(* IEC 61131-3 sources: kkh_knowHow_dgtt/tools/fmse/plc_lib, 31 files *)

(* ---- TYPES.st ---- *)
(*==================================================================================================================
  TYPES  -  enumerations and global constants of the FMSE device FB library
  ----------------------------------------------------------------------------------------------------------------
  Library   : FMSE device FB library (item 10A)              Version : 1.0.0 (2026-11-15)
  Rule      : tools/fmse/examples/item10a_examples.json  _rules.common, decisions D1 - D4
  Purpose   : one place for the state numbers (PackML item 5, device FBs), alarm classes and the time base.
              Load this file FIRST. Enumerations are used qualified (E_DriveState.FAULT); in CODESYS add
              the pragma attribute 'qualified_only', in TIA Portal use INT constants with the same values.
  Timing    : GC_CYCLE_MS = time base of the call counters of every FB. 100 = test bench (one call per
              100 ms tick). In the 10 ms main task set 10 - every time in ms stays the same.
  NOTICE    : ALL VALUES ARE EXAMPLES. Real PLC code is written, reviewed, tested and signed off by qualified
              people. Safety functions only in the F-program.
==================================================================================================================*)
TYPE
  E_AlarmClass : (NONE := 0, A := 1, B := 2, C := 3) INT;          (* decision D3 *)
  E_Reaction : (NONE := 0, ABORT := 1, HOLD := 2, WARNING := 3) INT;
  E_AlarmEvent : (NONE := 0, RAISE := 1, CLEAR := 2) INT;
  E_PackMLState : (UNDEFINED := 0, CLEARING := 1, STOPPED := 2, STARTING := 3, IDLE := 4, SUSPENDED := 5,
                   EXECUTE := 6, STOPPING := 7, ABORTING := 8, ABORTED := 9, HOLDING := 10, HELD := 11,
                   UNHOLDING := 12, SUSPENDING := 13, UNSUSPENDING := 14, RESETTING := 15, COMPLETING := 16,
                   COMPLETE := 17) INT;                             (* item 5, PackML / ISA-TR88 *)
  E_PackMLCmd : (NONE := 0, RESET := 1, START := 2, STOP := 3, HOLD := 4, UNHOLD := 5, SUSPEND := 6,
                 UNSUSPEND := 7, ABORT := 8, CLEAR := 9) INT;
  E_Mode : (UNDEFINED := 0, PRODUCTION := 1, MAINTENANCE := 2, MANUAL := 3) INT;
  E_DriveState : (NOT_READY := 0, READY := 1, RUNNING := 2, FAULT := 9) INT;
  E_MotorState : (STOPPED := 0, STARTING := 1, RUNNING := 2, STOPPING := 3, FAULT := 9) INT;
  E_HsStep : (IDLE := 0, REQUEST := 10, BUSY := 20, DONE := 30) INT;
  E_Quality : (GOOD := 0, UNCERTAIN := 1, BAD := 2) INT;             (* NAMUR NE 43 *)
  E_AiStatus : (OK := 0, FAULT_LOW := 1, UNDER_RANGE := 2, OVER_RANGE := 3, FAULT_HIGH := 4) INT;
END_TYPE

VAR_GLOBAL CONSTANT
  GC_CYCLE_MS : DINT := 100;                  (* time base of the call counters [ms] *)
  GC_N_MAX : DINT := 1000000;                 (* counters stop here (no overflow, 27 h at 100 ms) *)
  GC_BLINK_HALF_MS : DINT := 500;             (* half period of the 1 Hz blink [ms] *)
  GC_LIB_VERSION : WORD := 16#0100;           (* library version 1.0.0 *)
END_VAR

(* ---- F_CmdAllowed.st ---- *)
(*==================================================================================================================
  F_CmdAllowed  -  PackML command allowed in this state and mode? (item 5 tables)
  ----------------------------------------------------------------------------------------------------------------
  Library   : FMSE device FB library (item 10A)              Version : 1.0.0 (2026-11-15)
  Rule      : tools/fmse/examples/item10a_examples.json  _rules.FB_CmdIf
  Purpose   : TRUE when the command is in the mode table (1 Production: all 9, 2 Maintenance: without
              Suspend/Unsuspend, 3 Manual: Reset, Start, Stop, Abort, Clear) AND it is a transition of the
              state model: EDGES with the command label, Stop from every state except Stopped / Stopping /
              Aborting / Aborted / Clearing, Abort from every state except Aborting / Aborted.
  Interface :
    dir  name                type          default   meaning
    IN   iCmd                INT           -         command 1 Reset .. 9 Clear
    IN   iState              INT           -         PackML state 1 .. 17
    IN   iMode               INT           -         1 Production, 2 Maintenance, 3 Manual
  Alarms    : iAlarm = local code a ; Admin.AlarmNo = M*1000 + 10*i + a (decision D2), class per module (D3)
    none
  Timing    : Times are counted in calls: n * GC_CYCLE_MS >= t_ms (GC_CYCLE_MS = 100 ms = test bench, TYPES.st).
              In the 10 ms main task set GC_CYCLE_MS := 10 (same behaviour, 10 ms resolution) or replace a counter
              by a TON: ton(IN := <condition>, PT := T#2s); IF ton.Q THEN ... (one call later than the counter).
  Siemens   : SCL (TIA Portal): the same statements; local names are written with '#' (#xRst), the VAR section is
              VAR (STAT) of an FB with an instance DB, R_TRIG / TON are multi-instances, enumerations become INT
              constants (E_DriveState.FAULT -> 9), MIN / LIMIT exist, '16#0080' is written W#16#80 for a WORD.
  NOTICE    : ALL VALUES ARE EXAMPLES. Real PLC code is written, reviewed, tested and signed off by qualified
              people. Safety functions only in the F-program; this FB only reads F-copies and writes no F-signal.
==================================================================================================================*)
FUNCTION F_CmdAllowed : BOOL
VAR_INPUT  (* signals *)
  iCmd : INT;                               (* command 1 Reset .. 9 Clear *)
  iState : INT;                             (* PackML state 1 .. 17 *)
  iMode : INT;                              (* 1 Production, 2 Maintenance, 3 Manual *)
END_VAR
VAR  (* internal *)
  xInMode : BOOL;                           (* command allowed in the mode *)
END_VAR
F_CmdAllowed := FALSE;
CASE iMode OF
  E_Mode.PRODUCTION:
    xInMode := iCmd >= E_PackMLCmd.RESET AND iCmd <= E_PackMLCmd.CLEAR;
  E_Mode.MAINTENANCE:
    xInMode := (iCmd >= E_PackMLCmd.RESET AND iCmd <= E_PackMLCmd.UNHOLD) OR iCmd = E_PackMLCmd.ABORT
               OR iCmd = E_PackMLCmd.CLEAR;
  E_Mode.MANUAL:
    xInMode := (iCmd >= E_PackMLCmd.RESET AND iCmd <= E_PackMLCmd.STOP) OR iCmd = E_PackMLCmd.ABORT
               OR iCmd = E_PackMLCmd.CLEAR;
ELSE
  xInMode := FALSE;
END_CASE
IF NOT xInMode OR iState < E_PackMLState.CLEARING OR iState > E_PackMLState.COMPLETE THEN
  RETURN;
END_IF
CASE iCmd OF
  E_PackMLCmd.RESET:
    F_CmdAllowed := iState = E_PackMLState.STOPPED OR iState = E_PackMLState.COMPLETE;
  E_PackMLCmd.START:
    F_CmdAllowed := iState = E_PackMLState.IDLE;
  E_PackMLCmd.STOP:
    CASE iState OF
      E_PackMLState.CLEARING, E_PackMLState.STOPPED, E_PackMLState.STOPPING..E_PackMLState.ABORTED:
        F_CmdAllowed := FALSE;
    ELSE
      F_CmdAllowed := TRUE;
    END_CASE
  E_PackMLCmd.HOLD, E_PackMLCmd.SUSPEND:
    F_CmdAllowed := iState = E_PackMLState.EXECUTE;
  E_PackMLCmd.UNHOLD:
    F_CmdAllowed := iState = E_PackMLState.HELD;
  E_PackMLCmd.UNSUSPEND:
    F_CmdAllowed := iState = E_PackMLState.SUSPENDED;
  E_PackMLCmd.ABORT:
    F_CmdAllowed := iState <> E_PackMLState.ABORTING AND iState <> E_PackMLState.ABORTED;
  E_PackMLCmd.CLEAR:
    F_CmdAllowed := iState = E_PackMLState.ABORTED;
END_CASE
END_FUNCTION

(* ---- FB_AlarmMgr.st ---- *)
(*==================================================================================================================
  FB_AlarmMgr  -  module alarm manager: AlarmNo, WarningNo, class, reaction (D2 + D3)
  ----------------------------------------------------------------------------------------------------------------
  Library   : FMSE device FB library (item 10A)              Version : 1.0.0 (2026-11-15)
  Rule      : tools/fmse/examples/item10a_examples.json  _rules.alarm_manager
  Purpose   : Called once per alarm change (iEvent 1 = on, 2 = off; 0 = only evaluate) with the instance i, the
              local code a and the class of that alarm (class table generated from the library, item 10B).
              Admin.AlarmNo = best active class A/B alarm (A before B, earlier before later), Admin.WarningNo =
              earliest active class C, iAlarmClass for FB_SignalTower, iReaction for the PackML core.
  Interface :
    dir  name                type          default   meaning
    IN   iEvent              INT           -         0 none, 1 alarm on, 2 alarm off
    IN   iInst               INT           -         instance number i (0 = module level)
    IN   iCode               INT           -         local alarm code a (1 .. 9)
    IN   iClass              INT           -         class 1 A, 2 B, 3 C
    CFG  iModule             INT           2         module number M (M02 -> 2)
    OUT  iAlarmNo            INT           -         Admin.AlarmNo = M*1000 + 10*i + a
    OUT  iWarningNo          INT           -         Admin.WarningNo
    OUT  iAlarmClass         INT           -         0 none, 1 A, 2 B, 3 C
    OUT  iReaction           INT           -         0 none, 1 Abort, 2 Hold if Execute, 3 warning
    OUT  iActive             INT           -         number of active alarms
    OUT  xOverflow           BOOL          -         active list full
  Alarms    : iAlarm = local code a ; Admin.AlarmNo = M*1000 + 10*i + a (decision D2), class per module (D3)
    none
  Timing    : Times are counted in calls: n * GC_CYCLE_MS >= t_ms (GC_CYCLE_MS = 100 ms = test bench, TYPES.st).
              In the 10 ms main task set GC_CYCLE_MS := 10 (same behaviour, 10 ms resolution) or replace a counter
              by a TON: ton(IN := <condition>, PT := T#2s); IF ton.Q THEN ... (one call later than the counter).
  Siemens   : SCL (TIA Portal): the same statements; local names are written with '#' (#xRst), the VAR section is
              VAR (STAT) of an FB with an instance DB, R_TRIG / TON are multi-instances, enumerations become INT
              constants (E_DriveState.FAULT -> 9), MIN / LIMIT exist, '16#0080' is written W#16#80 for a WORD.
  NOTICE    : ALL VALUES ARE EXAMPLES. Real PLC code is written, reviewed, tested and signed off by qualified
              people. Safety functions only in the F-program; this FB only reads F-copies and writes no F-signal.
==================================================================================================================*)
FUNCTION_BLOCK FB_AlarmMgr
VAR_INPUT  (* signals *)
  iEvent : INT;                             (* 0 none, 1 alarm on, 2 alarm off *)
  iInst : INT;                              (* instance number i (0 = module level) *)
  iCode : INT;                              (* local alarm code a (1 .. 9) *)
  iClass : INT;                             (* class 1 A, 2 B, 3 C *)
END_VAR
VAR_INPUT  (* configuration (set once, defaults = example values) *)
  iModule : INT := 2;                       (* module number M (M02 -> 2) *)
END_VAR
VAR_OUTPUT  (* outputs *)
  iAlarmNo : INT;                           (* Admin.AlarmNo = M*1000 + 10*i + a *)
  iWarningNo : INT;                         (* Admin.WarningNo *)
  iAlarmClass : INT;                        (* 0 none, 1 A, 2 B, 3 C *)
  iReaction : INT;                          (* 0 none, 1 Abort, 2 Hold if Execute, 3 warning *)
  iActive : INT;                            (* number of active alarms *)
  xOverflow : BOOL;                         (* active list full *)
END_VAR
VAR CONSTANT  (* constants *)
  MAX_ACT : INT := 32;                      (* size of the active list *)
END_VAR
VAR  (* internal *)
  aiNo : ARRAY[1..MAX_ACT] OF INT;          (* active alarm numbers (0 = free) *)
  aiCls : ARRAY[1..MAX_ACT] OF INT;         (* class of each active alarm *)
  adiOrd : ARRAY[1..MAX_ACT] OF DINT;       (* activation order *)
  diOrder : DINT;                           (* activation counter *)
  iNo : INT;                                (* number of this event *)
  k : INT;                                  (* loop index *)
  iFound : INT;                             (* slot of iNo (0 = not active) *)
  iFree : INT;                              (* first free slot *)
  iBest : INT;                              (* slot of the best A/B alarm *)
  iBestW : INT;                             (* slot of the earliest warning *)
END_VAR
IF iEvent <> E_AlarmEvent.NONE THEN
  iNo := iModule * 1000 + 10 * iInst + iCode;
  iFound := 0;
  iFree := 0;
  FOR k := 1 TO MAX_ACT DO
    IF aiNo[k] = iNo AND iFound = 0 THEN
      iFound := k;
    END_IF
    IF aiNo[k] = 0 AND iFree = 0 THEN
      iFree := k;
    END_IF
  END_FOR
  IF iEvent = E_AlarmEvent.RAISE AND iFound = 0 THEN
    IF iFree > 0 THEN
      diOrder := diOrder + 1;
      aiNo[iFree] := iNo;
      aiCls[iFree] := iClass;
      adiOrd[iFree] := diOrder;
    ELSE
      xOverflow := TRUE;
    END_IF
  ELSIF iEvent = E_AlarmEvent.CLEAR AND iFound > 0 THEN
    aiNo[iFound] := 0;
    aiCls[iFound] := 0;
    adiOrd[iFound] := 0;
  END_IF
END_IF
(* evaluate: best class A/B alarm by (class, activation order), earliest class C warning *)
iBest := 0;
iBestW := 0;
iActive := 0;
FOR k := 1 TO MAX_ACT DO
  IF aiNo[k] <> 0 THEN
    iActive := iActive + 1;
    IF aiCls[k] = E_AlarmClass.A OR aiCls[k] = E_AlarmClass.B THEN
      IF iBest = 0 THEN
        iBest := k;
      ELSIF aiCls[k] < aiCls[iBest] OR (aiCls[k] = aiCls[iBest] AND adiOrd[k] < adiOrd[iBest]) THEN
        iBest := k;
      END_IF
    ELSIF aiCls[k] = E_AlarmClass.C THEN
      IF iBestW = 0 THEN
        iBestW := k;
      ELSIF adiOrd[k] < adiOrd[iBestW] THEN
        iBestW := k;
      END_IF
    END_IF
  END_IF
END_FOR
IF iBest > 0 THEN
  iAlarmNo := aiNo[iBest];
  iAlarmClass := aiCls[iBest];
ELSE
  iAlarmNo := 0;
  IF iBestW > 0 THEN
    iAlarmClass := E_AlarmClass.C;
  ELSE
    iAlarmClass := E_AlarmClass.NONE;
  END_IF
END_IF
IF iBestW > 0 THEN
  iWarningNo := aiNo[iBestW];
ELSE
  iWarningNo := 0;
END_IF
CASE iAlarmClass OF
  E_AlarmClass.A: iReaction := E_Reaction.ABORT;
  E_AlarmClass.B: iReaction := E_Reaction.HOLD;
  E_AlarmClass.C: iReaction := E_Reaction.WARNING;
ELSE
  iReaction := E_Reaction.NONE;
END_CASE
END_FUNCTION_BLOCK

(* ---- FB_AnalogIn.st ---- *)
(*==================================================================================================================
  FB_AnalogIn  -  4-20 mA analog input: scaling, NAMUR NE 43 quality, substitute value (item 9)
  ----------------------------------------------------------------------------------------------------------------
  Library   : FMSE device FB library (item 10A)              Version : 1.0.0 (2026-11-15)
  Rule      : tools/fmse/examples/item10a_examples.json  item9_examples.json _rules.analog
  Codegen   : item 8 pattern ANALOG_P, ANALOG_T -> st_codegen.py calls this FB (x<Signal> / q<Signal>)
  Purpose   : raw 0..27648 = 4..20 mA (Siemens-style card scaling - check yours). NE 43: <= 3.6 mA BAD (wire
              break), < 3.8 UNCERTAIN, <= 20.5 GOOD, < 21.0 UNCERTAIN, else BAD. rValue = clamped value for
              GOOD / UNCERTAIN, substitute rLo for BAD (the module must not use a BAD value).
  Interface :
    dir  name                type          default   meaning
    IN   iValue              INT           -         raw value of the card (AI)
    CFG  rLo                 REAL          0.0       value at 4 mA
    CFG  rHi                 REAL          10.0      value at 20 mA
    OUT  rMa                 REAL          -         current [mA]
    OUT  rValueLin           REAL          -         linear value (not clamped)
    OUT  rValue              REAL          -         value to use (clamped / substitute)
    OUT  iQuality            INT           -         0 GOOD, 1 UNCERTAIN, 2 BAD
    OUT  iStatus             INT           -         0 ok, 1 fault low, 2 under, 3 over, 4 fault high
    OUT  xGood               BOOL          -         quality GOOD
    OUT  iAlarm              INT           -         local alarm code (0 = none)
  Alarms    : iAlarm = local code a ; Admin.AlarmNo = M*1000 + 10*i + a (decision D2), class per module (D3)
    3  signal quality bad/uncertain (NAMUR NE 43)
  Timing    : Times are counted in calls: n * GC_CYCLE_MS >= t_ms (GC_CYCLE_MS = 100 ms = test bench, TYPES.st).
              In the 10 ms main task set GC_CYCLE_MS := 10 (same behaviour, 10 ms resolution) or replace a counter
              by a TON: ton(IN := <condition>, PT := T#2s); IF ton.Q THEN ... (one call later than the counter).
  Siemens   : SCL (TIA Portal): the same statements; local names are written with '#' (#xRst), the VAR section is
              VAR (STAT) of an FB with an instance DB, R_TRIG / TON are multi-instances, enumerations become INT
              constants (E_DriveState.FAULT -> 9), MIN / LIMIT exist, '16#0080' is written W#16#80 for a WORD.
  NOTICE    : ALL VALUES ARE EXAMPLES. Real PLC code is written, reviewed, tested and signed off by qualified
              people. Safety functions only in the F-program; this FB only reads F-copies and writes no F-signal.
==================================================================================================================*)
FUNCTION_BLOCK FB_AnalogIn
VAR_INPUT  (* signals *)
  iValue : INT;                             (* raw value of the card (AI) *)
END_VAR
VAR_INPUT  (* configuration (set once, defaults = example values) *)
  rLo : REAL := 0.0;                        (* value at 4 mA *)
  rHi : REAL := 10.0;                       (* value at 20 mA *)
END_VAR
VAR_OUTPUT  (* outputs *)
  rMa : REAL;                               (* current [mA] *)
  rValueLin : REAL;                         (* linear value (not clamped) *)
  rValue : REAL;                            (* value to use (clamped / substitute) *)
  iQuality : INT;                           (* 0 GOOD, 1 UNCERTAIN, 2 BAD *)
  iStatus : INT;                            (* 0 ok, 1 fault low, 2 under, 3 over, 4 fault high *)
  xGood : BOOL;                             (* quality GOOD *)
  iAlarm : INT;                             (* local alarm code (0 = none) *)
END_VAR
rMa := 4.0 + 16.0 * INT_TO_REAL(iValue) / 27648.0;
IF rMa <= 3.6 THEN
  iQuality := E_Quality.BAD;
  iStatus := E_AiStatus.FAULT_LOW;            (* wire break *)
ELSIF rMa < 3.8 THEN
  iQuality := E_Quality.UNCERTAIN;
  iStatus := E_AiStatus.UNDER_RANGE;
ELSIF rMa <= 20.5 THEN
  iQuality := E_Quality.GOOD;
  iStatus := E_AiStatus.OK;
ELSIF rMa < 21.0 THEN
  iQuality := E_Quality.UNCERTAIN;
  iStatus := E_AiStatus.OVER_RANGE;
ELSE
  iQuality := E_Quality.BAD;
  iStatus := E_AiStatus.FAULT_HIGH;
END_IF
rValueLin := rLo + (rHi - rLo) * (rMa - 4.0) / 16.0;
IF iQuality = E_Quality.BAD THEN
  rValue := rLo;                              (* substitute value *)
ELSE
  rValue := LIMIT(rLo, rValueLin, rHi);
END_IF
xGood := iQuality = E_Quality.GOOD;
IF xGood THEN
  iAlarm := 0;
ELSE
  iAlarm := 3;                                (* signal quality bad / uncertain *)
END_IF
END_FUNCTION_BLOCK

(* ---- FB_CmdIf.st ---- *)
(*==================================================================================================================
  FB_CmdIf  -  command interface of the module data block (4-phase echo, decision D1)
  ----------------------------------------------------------------------------------------------------------------
  Library   : FMSE device FB library (item 10A)              Version : 1.0.0 (2026-11-15)
  Rule      : tools/fmse/examples/item10a_examples.json  _rules.FB_CmdIf
  Purpose   : The cell controller writes CntrlCmd + sets CmdChangeRequest in ONE FC16 write. On the rising edge
              the module evaluates the command (F_CmdAllowed) -> CmdAck (Status.Bits bit8, iCmdExec one call
              for the PackML core) or CmdRej (bit9; the module sets Admin.WarningNo = M*1000 + 900 + command).
              The CC clears the request, then the module clears the echo. One writer per word, no command twice.
  Interface :
    dir  name                type          default   meaning
    IN   iCntrlCmd           INT           -         data block word CntrlCmd (written by the CC)
    IN   xCmdChangeRequest   BOOL          -         word 3 bit0 (written by the CC)
    IN   iState              INT           2         PackML state of the module
    IN   iMode               INT           1         mode of the module
    OUT  xCmdAck             BOOL          -         echo: accepted (Status.Bits bit8)
    OUT  xCmdRej             BOOL          -         echo: rejected (Status.Bits bit9)
    OUT  iCmdExec            INT           -         command to execute, one call (0 = none)
    OUT  iLastCmd            INT           -         last evaluated command
    OUT  iRejectCount        INT           -         rejected commands
  Alarms    : iAlarm = local code a ; Admin.AlarmNo = M*1000 + 10*i + a (decision D2), class per module (D3)
    none
  Timing    : Times are counted in calls: n * GC_CYCLE_MS >= t_ms (GC_CYCLE_MS = 100 ms = test bench, TYPES.st).
              In the 10 ms main task set GC_CYCLE_MS := 10 (same behaviour, 10 ms resolution) or replace a counter
              by a TON: ton(IN := <condition>, PT := T#2s); IF ton.Q THEN ... (one call later than the counter).
  Siemens   : SCL (TIA Portal): the same statements; local names are written with '#' (#xRst), the VAR section is
              VAR (STAT) of an FB with an instance DB, R_TRIG / TON are multi-instances, enumerations become INT
              constants (E_DriveState.FAULT -> 9), MIN / LIMIT exist, '16#0080' is written W#16#80 for a WORD.
  NOTICE    : ALL VALUES ARE EXAMPLES. Real PLC code is written, reviewed, tested and signed off by qualified
              people. Safety functions only in the F-program; this FB only reads F-copies and writes no F-signal.
==================================================================================================================*)
FUNCTION_BLOCK FB_CmdIf
VAR_INPUT  (* signals *)
  iCntrlCmd : INT;                          (* data block word CntrlCmd (written by the CC) *)
  xCmdChangeRequest : BOOL;                 (* word 3 bit0 (written by the CC) *)
  iState : INT := 2;                        (* PackML state of the module *)
  iMode : INT := 1;                         (* mode of the module *)
END_VAR
VAR_OUTPUT  (* outputs *)
  xCmdAck : BOOL;                           (* echo: accepted (Status.Bits bit8) *)
  xCmdRej : BOOL;                           (* echo: rejected (Status.Bits bit9) *)
  iCmdExec : INT;                           (* command to execute, one call (0 = none) *)
  iLastCmd : INT;                           (* last evaluated command *)
  iRejectCount : INT;                       (* rejected commands *)
END_VAR
VAR  (* internal *)
  rtReq : R_TRIG;                           (* edge of xCmdChangeRequest *)
END_VAR
rtReq(CLK := xCmdChangeRequest);
iCmdExec := 0;
IF rtReq.Q THEN
  iLastCmd := iCntrlCmd;
  IF F_CmdAllowed(iCmd := iCntrlCmd, iState := iState, iMode := iMode) THEN
    xCmdAck := TRUE;
    iCmdExec := iCntrlCmd;
  ELSE
    xCmdRej := TRUE;
    iRejectCount := iRejectCount + 1;
  END_IF
END_IF
IF NOT xCmdChangeRequest THEN                 (* phase 4: the CC has cleared the request *)
  xCmdAck := FALSE;
  xCmdRej := FALSE;
END_IF
END_FUNCTION_BLOCK

(* ---- FB_ContactorPair.st ---- *)
(*==================================================================================================================
  FB_ContactorPair  -  redundant contactor pair with EDM
  ----------------------------------------------------------------------------------------------------------------
  Library   : FMSE device FB library (item 10A)              Version : 1.0.0 (2026-11-15)
  Rule      : tools/fmse/examples/item10a_examples.json  _rules.fb_library (= FB_Edm, bInverted TRUE)
  Codegen   : item 8 pattern CONT_PAIR_EDM -> st_codegen.py calls this FB (x<Signal> / q<Signal>)
  Purpose   : Wrapper of FB_Edm with bInverted TRUE. The F-output Enable is written only by the F-program;
              xCmd is its read-only F-copy.
  Interface :
    dir  name                type          default   meaning
    IN   xCmd                BOOL          -         F-copy of the F-output Enable
    IN   xEDM                BOOL          TRUE      NC mirror contacts in series (DI), TRUE = open
    IN   xReset              BOOL          -         fault reset, rising edge
    CFG  tEdm_ms             DINT          300       feedback time [ms]
    OUT  xOn                 BOOL          -         output on and feedback ok
    OUT  xError              BOOL          -         error latched (see alarms)
    OUT  iAlarm              INT           -         local alarm code (0 = none)
  Alarms    : iAlarm = local code a ; Admin.AlarmNo = M*1000 + 10*i + a (decision D2), class per module (D3)
    1  feedback does not follow (welded / not switching)
  Timing    : Times are counted in calls: n * GC_CYCLE_MS >= t_ms (GC_CYCLE_MS = 100 ms = test bench, TYPES.st).
              In the 10 ms main task set GC_CYCLE_MS := 10 (same behaviour, 10 ms resolution) or replace a counter
              by a TON: ton(IN := <condition>, PT := T#2s); IF ton.Q THEN ... (one call later than the counter).
  Siemens   : SCL (TIA Portal): the same statements; local names are written with '#' (#xRst), the VAR section is
              VAR (STAT) of an FB with an instance DB, R_TRIG / TON are multi-instances, enumerations become INT
              constants (E_DriveState.FAULT -> 9), MIN / LIMIT exist, '16#0080' is written W#16#80 for a WORD.
  NOTICE    : ALL VALUES ARE EXAMPLES. Real PLC code is written, reviewed, tested and signed off by qualified
              people. Safety functions only in the F-program; this FB only reads F-copies and writes no F-signal.
==================================================================================================================*)
FUNCTION_BLOCK FB_ContactorPair
VAR_INPUT  (* signals *)
  xCmd : BOOL;                              (* F-copy of the F-output Enable *)
  xEDM : BOOL := TRUE;                      (* NC mirror contacts in series (DI), TRUE = open *)
  xReset : BOOL;                            (* fault reset, rising edge *)
END_VAR
VAR_INPUT  (* configuration (set once, defaults = example values) *)
  tEdm_ms : DINT := 300;                    (* feedback time [ms] *)
END_VAR
VAR_OUTPUT  (* outputs *)
  xOn : BOOL;                               (* output on and feedback ok *)
  xError : BOOL;                            (* error latched (see alarms) *)
  iAlarm : INT;                             (* local alarm code (0 = none) *)
END_VAR
VAR  (* internal *)
  fbEdm : FB_Edm;                           (* EDM *)
END_VAR
fbEdm(xCmd := xCmd, xFb := xEDM, xReset := xReset, tEdm_ms := tEdm_ms, bInverted := TRUE);
xOn := fbEdm.xOn;
xError := fbEdm.xError;
iAlarm := fbEdm.iAlarm;
END_FUNCTION_BLOCK

(* ---- FB_Door2Ch.st ---- *)
(*==================================================================================================================
  FB_Door2Ch  -  guard door switch (2 channels, no locking)
  ----------------------------------------------------------------------------------------------------------------
  Library   : FMSE device FB library (item 10A)              Version : 1.0.0 (2026-11-15)
  Rule      : tools/fmse/examples/item10a_examples.json  _rules.fb_library (= FB_Safe2Ch)
  Codegen   : item 8 pattern DOOR_2CH -> st_codegen.py calls this FB (x<Signal> / q<Signal>)
  Purpose   : Wrapper with the item-8 signal names: xClosed / xClosed2 -> FB_Safe2Ch xCh1 / xCh2.
              Diagnosis and HMI only - the safety function is in the F-program.
  Interface :
    dir  name                type          default   meaning
    IN   xClosed             BOOL          -         door closed channel 1 F-copy
    IN   xClosed2            BOOL          -         door closed channel 2 F-copy
    IN   xReset              BOOL          -         fault reset, rising edge
    CFG  tDisc_ms            DINT          500       discrepancy time [ms]
    OUT  xSafe               BOOL          -         closed / free and reset (FB_Safe2Ch.xOk)
    OUT  xResetReq           BOOL          -         waiting for a reset
    OUT  xDiscErr            BOOL          -         discrepancy latched
    OUT  iAlarm              INT           -         local alarm code (0 = none)
  Alarms    : iAlarm = local code a ; Admin.AlarmNo = M*1000 + 10*i + a (decision D2), class per module (D3)
    1  discrepancy
  Timing    : Times are counted in calls: n * GC_CYCLE_MS >= t_ms (GC_CYCLE_MS = 100 ms = test bench, TYPES.st).
              In the 10 ms main task set GC_CYCLE_MS := 10 (same behaviour, 10 ms resolution) or replace a counter
              by a TON: ton(IN := <condition>, PT := T#2s); IF ton.Q THEN ... (one call later than the counter).
  Siemens   : SCL (TIA Portal): the same statements; local names are written with '#' (#xRst), the VAR section is
              VAR (STAT) of an FB with an instance DB, R_TRIG / TON are multi-instances, enumerations become INT
              constants (E_DriveState.FAULT -> 9), MIN / LIMIT exist, '16#0080' is written W#16#80 for a WORD.
  NOTICE    : ALL VALUES ARE EXAMPLES. Real PLC code is written, reviewed, tested and signed off by qualified
              people. Safety functions only in the F-program; this FB only reads F-copies and writes no F-signal.
==================================================================================================================*)
FUNCTION_BLOCK FB_Door2Ch
VAR_INPUT  (* signals *)
  xClosed : BOOL;                           (* door closed channel 1 F-copy *)
  xClosed2 : BOOL;                          (* door closed channel 2 F-copy *)
  xReset : BOOL;                            (* fault reset, rising edge *)
END_VAR
VAR_INPUT  (* configuration (set once, defaults = example values) *)
  tDisc_ms : DINT := 500;                   (* discrepancy time [ms] *)
END_VAR
VAR_OUTPUT  (* outputs *)
  xSafe : BOOL;                             (* closed / free and reset (FB_Safe2Ch.xOk) *)
  xResetReq : BOOL;                         (* waiting for a reset *)
  xDiscErr : BOOL;                          (* discrepancy latched *)
  iAlarm : INT;                             (* local alarm code (0 = none) *)
END_VAR
VAR  (* internal *)
  fbCh : FB_Safe2Ch;                        (* 2-channel mirror *)
END_VAR
fbCh(xCh1 := xClosed, xCh2 := xClosed2, xReset := xReset, tDisc_ms := tDisc_ms);
xSafe := fbCh.xOk;
xResetReq := fbCh.xResetReq;
xDiscErr := fbCh.xDiscErr;
iAlarm := fbCh.iAlarm;
END_FUNCTION_BLOCK

(* ---- FB_DoorLock.st ---- *)
(*==================================================================================================================
  FB_DoorLock  -  guard locking: door + lock switch pairs, access request
  ----------------------------------------------------------------------------------------------------------------
  Library   : FMSE device FB library (item 10A)              Version : 1.0.0 (2026-11-15)
  Rule      : tools/fmse/examples/item10a_examples.json  _rules.FB_DoorLock
  Codegen   : item 8 pattern DOOR_LOCK -> st_codegen.py calls this FB (x<Signal> / q<Signal>)
  Purpose   : Item 7/8 DOOR_LOCK: discrepancy of the door pair and of the lock pair, locked-but-not-closed
              (tongue missing / manipulation), access request to the F-program (unlock after standstill), the
              request ends when the door was opened and closed again. Errors are latched (module reset, part B).
  Interface :
    dir  name                type          default   meaning
    IN   xClosed             BOOL          TRUE      door closed, channel 1 (DI)
    IN   xClosed2            BOOL          TRUE      door closed, channel 2 (DI)
    IN   xLocked             BOOL          TRUE      tongue locked, channel 1 (DI)
    IN   xLocked2            BOOL          TRUE      tongue locked, channel 2 (DI)
    IN   xRequest            BOOL          -         access request button, rising edge
    CFG  tDisc_ms            DINT          500       discrepancy time [ms]
    OUT  xClosedOk           BOOL          -         door closed (both)
    OUT  xLockedOk           BOOL          -         locked (both)
    OUT  xUnlockReq          BOOL          -         unlock request to the F-program
    OUT  xError              BOOL          -         error latched (see alarms)
    OUT  iAlarm              INT           -         local alarm code (0 = none)
  Alarms    : iAlarm = local code a ; Admin.AlarmNo = M*1000 + 10*i + a (decision D2), class per module (D3)
    1  door switch discrepancy
    2  lock switch discrepancy
    3  locked but not closed (tongue missing / manipulation)
  Timing    : Times are counted in calls: n * GC_CYCLE_MS >= t_ms (GC_CYCLE_MS = 100 ms = test bench, TYPES.st).
              In the 10 ms main task set GC_CYCLE_MS := 10 (same behaviour, 10 ms resolution) or replace a counter
              by a TON: ton(IN := <condition>, PT := T#2s); IF ton.Q THEN ... (one call later than the counter).
  Siemens   : SCL (TIA Portal): the same statements; local names are written with '#' (#xRst), the VAR section is
              VAR (STAT) of an FB with an instance DB, R_TRIG / TON are multi-instances, enumerations become INT
              constants (E_DriveState.FAULT -> 9), MIN / LIMIT exist, '16#0080' is written W#16#80 for a WORD.
  NOTICE    : ALL VALUES ARE EXAMPLES. Real PLC code is written, reviewed, tested and signed off by qualified
              people. Safety functions only in the F-program; this FB only reads F-copies and writes no F-signal.
==================================================================================================================*)
FUNCTION_BLOCK FB_DoorLock
VAR_INPUT  (* signals *)
  xClosed : BOOL := TRUE;                   (* door closed, channel 1 (DI) *)
  xClosed2 : BOOL := TRUE;                  (* door closed, channel 2 (DI) *)
  xLocked : BOOL := TRUE;                   (* tongue locked, channel 1 (DI) *)
  xLocked2 : BOOL := TRUE;                  (* tongue locked, channel 2 (DI) *)
  xRequest : BOOL;                          (* access request button, rising edge *)
END_VAR
VAR_INPUT  (* configuration (set once, defaults = example values) *)
  tDisc_ms : DINT := 500;                   (* discrepancy time [ms] *)
END_VAR
VAR_OUTPUT  (* outputs *)
  xClosedOk : BOOL;                         (* door closed (both) *)
  xLockedOk : BOOL;                         (* locked (both) *)
  xUnlockReq : BOOL;                        (* unlock request to the F-program *)
  xError : BOOL;                            (* error latched (see alarms) *)
  iAlarm : INT;                             (* local alarm code (0 = none) *)
END_VAR
VAR  (* internal *)
  rtReq : R_TRIG;                           (* edge of xRequest *)
  xC : BOOL;                                (* closed (both) *)
  xL : BOOL;                                (* locked (both) *)
  nC : DINT;                                (* door pair discrepancy calls *)
  nL : DINT;                                (* lock pair discrepancy calls *)
  xWasOpen : BOOL;                          (* door was open during the request *)
END_VAR
rtReq(CLK := xRequest);
xC := xClosed AND xClosed2;
xL := xLocked AND xLocked2;
IF xClosed <> xClosed2 THEN
  nC := MIN(nC + 1, GC_N_MAX);
ELSE
  nC := 0;
END_IF
IF xLocked <> xLocked2 THEN
  nL := MIN(nL + 1, GC_N_MAX);
ELSE
  nL := 0;
END_IF
IF nC * GC_CYCLE_MS >= tDisc_ms THEN
  xError := TRUE;
  iAlarm := 1;                                (* door switch discrepancy *)
ELSIF nL * GC_CYCLE_MS >= tDisc_ms THEN
  xError := TRUE;
  iAlarm := 2;                                (* lock switch discrepancy *)
END_IF
IF xL AND NOT xC AND NOT xError THEN
  xError := TRUE;
  iAlarm := 3;                                (* locked but not closed *)
END_IF
IF rtReq.Q AND xC AND xL THEN
  xUnlockReq := TRUE;
END_IF
IF NOT xClosed AND NOT xClosed2 THEN
  xWasOpen := TRUE;
END_IF
IF xUnlockReq AND xWasOpen AND xC THEN
  xUnlockReq := FALSE;                        (* opened and closed again: request done *)
  xWasOpen := FALSE;
END_IF
xClosedOk := xC;
xLockedOk := xL;
END_FUNCTION_BLOCK

(* ---- FB_DriveSto.st ---- *)
(*==================================================================================================================
  FB_DriveSto  -  frequency inverter with safe torque off (STO)
  ----------------------------------------------------------------------------------------------------------------
  Library   : FMSE device FB library (item 10A)              Version : 1.0.0 (2026-11-15)
  Rule      : tools/fmse/examples/item10a_examples.json  _rules.FB_DriveSto
  Codegen   : item 8 pattern VFD_STO -> st_codegen.py calls this FB (x<Signal> / q<Signal>)
  Purpose   : State machine of a drive whose STO is switched by the F-program (the standard program reads the
              F-copy xSto). STO is a normal safety stop, not a drive fault. wCtrl = control word over the bus.
  Interface :
    dir  name                type          default   meaning
    IN   xReady              BOOL          -         drive ready (DI)
    IN   xFault              BOOL          -         drive fault (DI)
    IN   xSto                BOOL          TRUE      F-copy: TRUE = torque off
    IN   xCmdRun             BOOL          -         run command from the sequence
    IN   xReset              BOOL          -         fault reset, rising edge
    OUT  wCtrl               WORD          -         bit0 enable, bit1 run, bit7 fault ack
    OUT  iState              INT           -         0 not ready, 1 ready, 2 running, 9 fault
    OUT  xWarn               BOOL          -         run requested while torque off
    OUT  xError              BOOL          -         error latched (see alarms)
    OUT  iAlarm              INT           -         local alarm code (0 = none)
  Alarms    : iAlarm = local code a ; Admin.AlarmNo = M*1000 + 10*i + a (decision D2), class per module (D3)
    1  drive fault
    3  ready lost while running
  Timing    : Times are counted in calls: n * GC_CYCLE_MS >= t_ms (GC_CYCLE_MS = 100 ms = test bench, TYPES.st).
              In the 10 ms main task set GC_CYCLE_MS := 10 (same behaviour, 10 ms resolution) or replace a counter
              by a TON: ton(IN := <condition>, PT := T#2s); IF ton.Q THEN ... (one call later than the counter).
  Siemens   : SCL (TIA Portal): the same statements; local names are written with '#' (#xRst), the VAR section is
              VAR (STAT) of an FB with an instance DB, R_TRIG / TON are multi-instances, enumerations become INT
              constants (E_DriveState.FAULT -> 9), MIN / LIMIT exist, '16#0080' is written W#16#80 for a WORD.
  NOTICE    : ALL VALUES ARE EXAMPLES. Real PLC code is written, reviewed, tested and signed off by qualified
              people. Safety functions only in the F-program; this FB only reads F-copies and writes no F-signal.
==================================================================================================================*)
FUNCTION_BLOCK FB_DriveSto
VAR_INPUT  (* signals *)
  xReady : BOOL;                            (* drive ready (DI) *)
  xFault : BOOL;                            (* drive fault (DI) *)
  xSto : BOOL := TRUE;                      (* F-copy: TRUE = torque off *)
  xCmdRun : BOOL;                           (* run command from the sequence *)
  xReset : BOOL;                            (* fault reset, rising edge *)
END_VAR
VAR_OUTPUT  (* outputs *)
  wCtrl : WORD;                             (* bit0 enable, bit1 run, bit7 fault ack *)
  iState : INT;                             (* 0 not ready, 1 ready, 2 running, 9 fault *)
  xWarn : BOOL;                             (* run requested while torque off *)
  xError : BOOL;                            (* error latched (see alarms) *)
  iAlarm : INT;                             (* local alarm code (0 = none) *)
END_VAR
VAR  (* internal *)
  rtReset : R_TRIG;                         (* edge of xReset *)
  xRst : BOOL;                              (* reset pulse *)
  xAck : BOOL;                              (* fault acknowledge, one call *)
END_VAR
rtReset(CLK := xReset);
xRst := rtReset.Q;
xAck := FALSE;
IF xFault AND iState <> E_DriveState.FAULT THEN
  iState := E_DriveState.FAULT;
  iAlarm := 1;                                (* drive fault *)
ELSE
  CASE iState OF                              (* one transition per call *)
    E_DriveState.NOT_READY:
      IF xReady AND NOT xSto THEN
        iState := E_DriveState.READY;
      END_IF
    E_DriveState.READY:
      IF xSto OR NOT xReady THEN
        iState := E_DriveState.NOT_READY;
      ELSIF xCmdRun THEN
        iState := E_DriveState.RUNNING;
      END_IF
    E_DriveState.RUNNING:
      IF xSto THEN
        iState := E_DriveState.NOT_READY;     (* STO = normal safety stop *)
      ELSIF NOT xReady THEN
        iState := E_DriveState.FAULT;
        iAlarm := 3;                          (* ready lost while running *)
      ELSIF NOT xCmdRun THEN
        iState := E_DriveState.READY;
      END_IF
    E_DriveState.FAULT:
      IF xRst AND NOT xFault THEN
        iState := E_DriveState.NOT_READY;
        iAlarm := 0;
        xAck := TRUE;
      END_IF
  END_CASE
END_IF
xError := iState = E_DriveState.FAULT;
xWarn := xCmdRun AND xSto;
wCtrl := 16#0000;
IF NOT xSto THEN
  wCtrl := wCtrl OR 16#0001;                  (* bit0 ON / enable *)
END_IF
IF iState = E_DriveState.RUNNING THEN
  wCtrl := wCtrl OR 16#0002;                  (* bit1 RUN *)
END_IF
IF xAck THEN
  wCtrl := wCtrl OR 16#0080;                  (* bit7 fault acknowledge *)
END_IF
END_FUNCTION_BLOCK

(* ---- FB_Edm.st ---- *)
(*==================================================================================================================
  FB_Edm  -  external device monitoring (EDM) of a safety output
  ----------------------------------------------------------------------------------------------------------------
  Library   : FMSE device FB library (item 10A)              Version : 1.0.0 (2026-11-15)
  Rule      : tools/fmse/examples/item10a_examples.json  _rules.FB_Edm
  Purpose   : Checks that the feedback of a safety output follows its command: NC mirror contacts of
              contactors (bInverted TRUE: feedback TRUE when OPEN) or the position switch of a safety valve
              (bInverted FALSE). Base of FB_ZoneOut, FB_ContactorPair and FB_SafeValve.
  Interface :
    dir  name                type          default   meaning
    IN   xCmd                BOOL          -         F-copy of the F-output (read only)
    IN   xFb                 BOOL          TRUE      feedback (DI)
    IN   xReset              BOOL          -         fault reset, rising edge
    CFG  tEdm_ms             DINT          300       feedback time [ms]
    CFG  bInverted           BOOL          TRUE      TRUE = NC mirror contact
    OUT  xOn                 BOOL          -         output on and feedback ok
    OUT  xError              BOOL          -         error latched (see alarms)
    OUT  iAlarm              INT           -         local alarm code (0 = none)
  Alarms    : iAlarm = local code a ; Admin.AlarmNo = M*1000 + 10*i + a (decision D2), class per module (D3)
    1  feedback does not follow (welded / not switching)
  Timing    : Times are counted in calls: n * GC_CYCLE_MS >= t_ms (GC_CYCLE_MS = 100 ms = test bench, TYPES.st).
              In the 10 ms main task set GC_CYCLE_MS := 10 (same behaviour, 10 ms resolution) or replace a counter
              by a TON: ton(IN := <condition>, PT := T#2s); IF ton.Q THEN ... (one call later than the counter).
  Siemens   : SCL (TIA Portal): the same statements; local names are written with '#' (#xRst), the VAR section is
              VAR (STAT) of an FB with an instance DB, R_TRIG / TON are multi-instances, enumerations become INT
              constants (E_DriveState.FAULT -> 9), MIN / LIMIT exist, '16#0080' is written W#16#80 for a WORD.
  NOTICE    : ALL VALUES ARE EXAMPLES. Real PLC code is written, reviewed, tested and signed off by qualified
              people. Safety functions only in the F-program; this FB only reads F-copies and writes no F-signal.
==================================================================================================================*)
FUNCTION_BLOCK FB_Edm
VAR_INPUT  (* signals *)
  xCmd : BOOL;                              (* F-copy of the F-output (read only) *)
  xFb : BOOL := TRUE;                       (* feedback (DI) *)
  xReset : BOOL;                            (* fault reset, rising edge *)
END_VAR
VAR_INPUT  (* configuration (set once, defaults = example values) *)
  tEdm_ms : DINT := 300;                    (* feedback time [ms] *)
  bInverted : BOOL := TRUE;                 (* TRUE = NC mirror contact *)
END_VAR
VAR_OUTPUT  (* outputs *)
  xOn : BOOL;                               (* output on and feedback ok *)
  xError : BOOL;                            (* error latched (see alarms) *)
  iAlarm : INT;                             (* local alarm code (0 = none) *)
END_VAR
VAR  (* internal *)
  rtReset : R_TRIG;                         (* edge of xReset *)
  xExp : BOOL;                              (* expected feedback *)
  xFbOk : BOOL;                             (* feedback = expected *)
  n : DINT;                                 (* calls with wrong feedback *)
END_VAR
rtReset(CLK := xReset);
IF bInverted THEN
  xExp := NOT xCmd;
ELSE
  xExp := xCmd;
END_IF
xFbOk := xFb = xExp;
IF NOT xFbOk THEN
  n := MIN(n + 1, GC_N_MAX);
ELSE
  n := 0;
END_IF
IF xError AND rtReset.Q AND xFbOk THEN
  xError := FALSE;
  iAlarm := 0;
END_IF
IF NOT xError AND n * GC_CYCLE_MS >= tEdm_ms THEN
  xError := TRUE;
  iAlarm := 1;                                (* feedback does not follow *)
END_IF
xOn := xCmd AND xFbOk AND NOT xError;
END_FUNCTION_BLOCK

(* ---- FB_EnableSwitch.st ---- *)
(*==================================================================================================================
  FB_EnableSwitch  -  3-position enabling switch (2 channels)
  ----------------------------------------------------------------------------------------------------------------
  Library   : FMSE device FB library (item 10A)              Version : 1.0.0 (2026-11-15)
  Rule      : tools/fmse/examples/item10a_examples.json  _rules.fb_library (= FB_Safe2Ch)
  Codegen   : item 8 pattern ENABLE -> st_codegen.py calls this FB (x<Signal> / q<Signal>)
  Purpose   : Wrapper with the item-8 signal names: xOk / xOk2 -> FB_Safe2Ch xCh1 / xCh2.
              Diagnosis and HMI only - the safety function is in the F-program.
  Interface :
    dir  name                type          default   meaning
    IN   xOk                 BOOL          -         enabling channel 1 F-copy (TRUE = enabled)
    IN   xOk2                BOOL          -         enabling channel 2 F-copy (TRUE = enabled)
    IN   xReset              BOOL          -         fault reset, rising edge
    CFG  tDisc_ms            DINT          500       discrepancy time [ms]
    OUT  xSafe               BOOL          -         closed / free and reset (FB_Safe2Ch.xOk)
    OUT  xResetReq           BOOL          -         waiting for a reset
    OUT  xDiscErr            BOOL          -         discrepancy latched
    OUT  iAlarm              INT           -         local alarm code (0 = none)
  Alarms    : iAlarm = local code a ; Admin.AlarmNo = M*1000 + 10*i + a (decision D2), class per module (D3)
    1  discrepancy
  Timing    : Times are counted in calls: n * GC_CYCLE_MS >= t_ms (GC_CYCLE_MS = 100 ms = test bench, TYPES.st).
              In the 10 ms main task set GC_CYCLE_MS := 10 (same behaviour, 10 ms resolution) or replace a counter
              by a TON: ton(IN := <condition>, PT := T#2s); IF ton.Q THEN ... (one call later than the counter).
  Siemens   : SCL (TIA Portal): the same statements; local names are written with '#' (#xRst), the VAR section is
              VAR (STAT) of an FB with an instance DB, R_TRIG / TON are multi-instances, enumerations become INT
              constants (E_DriveState.FAULT -> 9), MIN / LIMIT exist, '16#0080' is written W#16#80 for a WORD.
  NOTICE    : ALL VALUES ARE EXAMPLES. Real PLC code is written, reviewed, tested and signed off by qualified
              people. Safety functions only in the F-program; this FB only reads F-copies and writes no F-signal.
==================================================================================================================*)
FUNCTION_BLOCK FB_EnableSwitch
VAR_INPUT  (* signals *)
  xOk : BOOL;                               (* enabling channel 1 F-copy (TRUE = enabled) *)
  xOk2 : BOOL;                              (* enabling channel 2 F-copy (TRUE = enabled) *)
  xReset : BOOL;                            (* fault reset, rising edge *)
END_VAR
VAR_INPUT  (* configuration (set once, defaults = example values) *)
  tDisc_ms : DINT := 500;                   (* discrepancy time [ms] *)
END_VAR
VAR_OUTPUT  (* outputs *)
  xSafe : BOOL;                             (* closed / free and reset (FB_Safe2Ch.xOk) *)
  xResetReq : BOOL;                         (* waiting for a reset *)
  xDiscErr : BOOL;                          (* discrepancy latched *)
  iAlarm : INT;                             (* local alarm code (0 = none) *)
END_VAR
VAR  (* internal *)
  fbCh : FB_Safe2Ch;                        (* 2-channel mirror *)
END_VAR
fbCh(xCh1 := xOk, xCh2 := xOk2, xReset := xReset, tDisc_ms := tDisc_ms);
xSafe := fbCh.xOk;
xResetReq := fbCh.xResetReq;
xDiscErr := fbCh.xDiscErr;
iAlarm := fbCh.iAlarm;
END_FUNCTION_BLOCK

(* ---- FB_Estop.st ---- *)
(*==================================================================================================================
  FB_Estop  -  emergency stop button (2 channels)
  ----------------------------------------------------------------------------------------------------------------
  Library   : FMSE device FB library (item 10A)              Version : 1.0.0 (2026-11-15)
  Rule      : tools/fmse/examples/item10a_examples.json  _rules.fb_library (= FB_Safe2Ch)
  Codegen   : item 8 pattern ESTOP -> st_codegen.py calls this FB (x<Signal> / q<Signal>)
  Purpose   : Wrapper with the item-8 signal names: xOk / xOk2 -> FB_Safe2Ch xCh1 / xCh2.
              Diagnosis and HMI only - the safety function is in the F-program.
  Interface :
    dir  name                type          default   meaning
    IN   xOk                 BOOL          -         e-stop channel 1 F-copy (TRUE = not pressed)
    IN   xOk2                BOOL          -         e-stop channel 2 F-copy (TRUE = not pressed)
    IN   xReset              BOOL          -         fault reset, rising edge
    CFG  tDisc_ms            DINT          500       discrepancy time [ms]
    OUT  xSafe               BOOL          -         closed / free and reset (FB_Safe2Ch.xOk)
    OUT  xResetReq           BOOL          -         waiting for a reset
    OUT  xDiscErr            BOOL          -         discrepancy latched
    OUT  iAlarm              INT           -         local alarm code (0 = none)
  Alarms    : iAlarm = local code a ; Admin.AlarmNo = M*1000 + 10*i + a (decision D2), class per module (D3)
    1  discrepancy
  Timing    : Times are counted in calls: n * GC_CYCLE_MS >= t_ms (GC_CYCLE_MS = 100 ms = test bench, TYPES.st).
              In the 10 ms main task set GC_CYCLE_MS := 10 (same behaviour, 10 ms resolution) or replace a counter
              by a TON: ton(IN := <condition>, PT := T#2s); IF ton.Q THEN ... (one call later than the counter).
  Siemens   : SCL (TIA Portal): the same statements; local names are written with '#' (#xRst), the VAR section is
              VAR (STAT) of an FB with an instance DB, R_TRIG / TON are multi-instances, enumerations become INT
              constants (E_DriveState.FAULT -> 9), MIN / LIMIT exist, '16#0080' is written W#16#80 for a WORD.
  NOTICE    : ALL VALUES ARE EXAMPLES. Real PLC code is written, reviewed, tested and signed off by qualified
              people. Safety functions only in the F-program; this FB only reads F-copies and writes no F-signal.
==================================================================================================================*)
FUNCTION_BLOCK FB_Estop
VAR_INPUT  (* signals *)
  xOk : BOOL;                               (* e-stop channel 1 F-copy (TRUE = not pressed) *)
  xOk2 : BOOL;                              (* e-stop channel 2 F-copy (TRUE = not pressed) *)
  xReset : BOOL;                            (* fault reset, rising edge *)
END_VAR
VAR_INPUT  (* configuration (set once, defaults = example values) *)
  tDisc_ms : DINT := 500;                   (* discrepancy time [ms] *)
END_VAR
VAR_OUTPUT  (* outputs *)
  xSafe : BOOL;                             (* closed / free and reset (FB_Safe2Ch.xOk) *)
  xResetReq : BOOL;                         (* waiting for a reset *)
  xDiscErr : BOOL;                          (* discrepancy latched *)
  iAlarm : INT;                             (* local alarm code (0 = none) *)
END_VAR
VAR  (* internal *)
  fbCh : FB_Safe2Ch;                        (* 2-channel mirror *)
END_VAR
fbCh(xCh1 := xOk, xCh2 := xOk2, xReset := xReset, tDisc_ms := tDisc_ms);
xSafe := fbCh.xOk;
xResetReq := fbCh.xResetReq;
xDiscErr := fbCh.xDiscErr;
iAlarm := fbCh.iAlarm;
END_FUNCTION_BLOCK

(* ---- FB_Feeder.st ---- *)
(*==================================================================================================================
  FB_Feeder  -  external feeder / breaker monitoring
  ----------------------------------------------------------------------------------------------------------------
  Library   : FMSE device FB library (item 10A)              Version : 1.0.0 (2026-11-15)
  Rule      : tools/fmse/examples/item10a_examples.json  _rules.FB_Feeder
  Codegen   : item 8 pattern FEEDER_EXT -> st_codegen.py calls this FB (x<Signal> / q<Signal>)
  Purpose   : Auxiliary contact of a feeder breaker: alarm after tDelay_ms without supply (not latched).
  Interface :
    dir  name                type          default   meaning
    IN   xSupplyOn           BOOL          TRUE      breaker auxiliary contact (DI)
    CFG  tDelay_ms           DINT          200       alarm delay [ms]
    OUT  xOk                 BOOL          -         supply on
    OUT  iAlarm              INT           -         local alarm code (0 = none)
  Alarms    : iAlarm = local code a ; Admin.AlarmNo = M*1000 + 10*i + a (decision D2), class per module (D3)
    1  feeder breaker off
  Timing    : Times are counted in calls: n * GC_CYCLE_MS >= t_ms (GC_CYCLE_MS = 100 ms = test bench, TYPES.st).
              In the 10 ms main task set GC_CYCLE_MS := 10 (same behaviour, 10 ms resolution) or replace a counter
              by a TON: ton(IN := <condition>, PT := T#2s); IF ton.Q THEN ... (one call later than the counter).
  Siemens   : SCL (TIA Portal): the same statements; local names are written with '#' (#xRst), the VAR section is
              VAR (STAT) of an FB with an instance DB, R_TRIG / TON are multi-instances, enumerations become INT
              constants (E_DriveState.FAULT -> 9), MIN / LIMIT exist, '16#0080' is written W#16#80 for a WORD.
  NOTICE    : ALL VALUES ARE EXAMPLES. Real PLC code is written, reviewed, tested and signed off by qualified
              people. Safety functions only in the F-program; this FB only reads F-copies and writes no F-signal.
==================================================================================================================*)
FUNCTION_BLOCK FB_Feeder
VAR_INPUT  (* signals *)
  xSupplyOn : BOOL := TRUE;                 (* breaker auxiliary contact (DI) *)
END_VAR
VAR_INPUT  (* configuration (set once, defaults = example values) *)
  tDelay_ms : DINT := 200;                  (* alarm delay [ms] *)
END_VAR
VAR_OUTPUT  (* outputs *)
  xOk : BOOL;                               (* supply on *)
  iAlarm : INT;                             (* local alarm code (0 = none) *)
END_VAR
VAR  (* internal *)
  n : DINT;                                 (* calls without supply *)
END_VAR
IF NOT xSupplyOn THEN
  n := MIN(n + 1, GC_N_MAX);
ELSE
  n := 0;
END_IF
xOk := xSupplyOn;
IF n * GC_CYCLE_MS >= tDelay_ms THEN
  iAlarm := 1;                                (* feeder breaker off *)
ELSE
  iAlarm := 0;
END_IF
END_FUNCTION_BLOCK

(* ---- FB_HandshakeHw.st ---- *)
(*==================================================================================================================
  FB_HandshakeHw  -  requester side of the hard-wired 4-phase handshake
  ----------------------------------------------------------------------------------------------------------------
  Library   : FMSE device FB library (item 10A)              Version : 1.0.0 (2026-11-15)
  Rule      : tools/fmse/examples/item10a_examples.json  _rules.FB_HandshakeHw
  Codegen   : item 8 pattern HANDSHAKE_HW -> st_codegen.py calls this FB (x<Signal> / q<Signal>)
  Purpose   : Item 8 HANDSHAKE_HW / item 6 logic: Request + Enable -> partner Busy -> partner Done -> Ack ->
              partner removes Done -> finished (xDoneOut one call). Time-outs per phase, partner fault, reset.
  Interface :
    dir  name                type          default   meaning
    IN   xReady              BOOL          -         partner ready (DI)
    IN   xBusy               BOOL          -         partner busy (DI)
    IN   xDone               BOOL          -         partner done (DI)
    IN   xFault              BOOL          -         partner fault (DI)
    IN   xStart              BOOL          -         start a job (sequence)
    IN   xReset              BOOL          -         fault reset, rising edge
    CFG  tHs_ms              DINT          2000      handshake phase time-out [ms]
    CFG  tJob_ms             DINT          10000     job time-out [ms]
    OUT  qRequest            BOOL          -         request to the partner (DO)
    OUT  qAck                BOOL          -         acknowledge to the partner (DO)
    OUT  qEnable             BOOL          -         enable to the partner (DO)
    OUT  qReset              BOOL          -         fault reset to the partner, one call (DO)
    OUT  iStep               INT           -         0 idle, 10 request, 20 busy, 30 done
    OUT  xDoneOut            BOOL          -         job finished, one call
    OUT  xError              BOOL          -         error latched (see alarms)
    OUT  iAlarm              INT           -         local alarm code (0 = none)
  Alarms    : iAlarm = local code a ; Admin.AlarmNo = M*1000 + 10*i + a (decision D2), class per module (D3)
    1  partner did not start (busy missing)
    2  job time-out
    3  done not removed
    4  partner fault
  Timing    : Times are counted in calls: n * GC_CYCLE_MS >= t_ms (GC_CYCLE_MS = 100 ms = test bench, TYPES.st).
              In the 10 ms main task set GC_CYCLE_MS := 10 (same behaviour, 10 ms resolution) or replace a counter
              by a TON: ton(IN := <condition>, PT := T#2s); IF ton.Q THEN ... (one call later than the counter).
  Siemens   : SCL (TIA Portal): the same statements; local names are written with '#' (#xRst), the VAR section is
              VAR (STAT) of an FB with an instance DB, R_TRIG / TON are multi-instances, enumerations become INT
              constants (E_DriveState.FAULT -> 9), MIN / LIMIT exist, '16#0080' is written W#16#80 for a WORD.
  NOTICE    : ALL VALUES ARE EXAMPLES. Real PLC code is written, reviewed, tested and signed off by qualified
              people. Safety functions only in the F-program; this FB only reads F-copies and writes no F-signal.
==================================================================================================================*)
FUNCTION_BLOCK FB_HandshakeHw
VAR_INPUT  (* signals *)
  xReady : BOOL;                            (* partner ready (DI) *)
  xBusy : BOOL;                             (* partner busy (DI) *)
  xDone : BOOL;                             (* partner done (DI) *)
  xFault : BOOL;                            (* partner fault (DI) *)
  xStart : BOOL;                            (* start a job (sequence) *)
  xReset : BOOL;                            (* fault reset, rising edge *)
END_VAR
VAR_INPUT  (* configuration (set once, defaults = example values) *)
  tHs_ms : DINT := 2000;                    (* handshake phase time-out [ms] *)
  tJob_ms : DINT := 10000;                  (* job time-out [ms] *)
END_VAR
VAR_OUTPUT  (* outputs *)
  qRequest : BOOL;                          (* request to the partner (DO) *)
  qAck : BOOL;                              (* acknowledge to the partner (DO) *)
  qEnable : BOOL;                           (* enable to the partner (DO) *)
  qReset : BOOL;                            (* fault reset to the partner, one call (DO) *)
  iStep : INT;                              (* 0 idle, 10 request, 20 busy, 30 done *)
  xDoneOut : BOOL;                          (* job finished, one call *)
  xError : BOOL;                            (* error latched (see alarms) *)
  iAlarm : INT;                             (* local alarm code (0 = none) *)
END_VAR
VAR  (* internal *)
  rtReset : R_TRIG;                         (* edge of xReset *)
  xRst : BOOL;                              (* reset pulse *)
  n : DINT;                                 (* calls in the step *)
END_VAR
rtReset(CLK := xReset);
xRst := rtReset.Q;
qReset := xRst;
xDoneOut := FALSE;
IF xError THEN
  IF xRst AND NOT xFault THEN
    xError := FALSE;
    iAlarm := 0;
    iStep := E_HsStep.IDLE;
  END_IF
ELSIF xFault AND iStep <> E_HsStep.IDLE THEN
  xError := TRUE;
  iAlarm := 4;                                (* partner fault *)
ELSE
  CASE iStep OF
    E_HsStep.IDLE:
      IF xStart AND xReady THEN
        iStep := E_HsStep.REQUEST;
        n := 0;
      END_IF
    E_HsStep.REQUEST:
      n := MIN(n + 1, GC_N_MAX);
      IF xBusy THEN
        iStep := E_HsStep.BUSY;
        n := 0;
      ELSIF n * GC_CYCLE_MS >= tHs_ms THEN
        xError := TRUE;
        iAlarm := 1;                          (* partner did not start *)
      END_IF
    E_HsStep.BUSY:
      n := MIN(n + 1, GC_N_MAX);
      IF xDone THEN
        iStep := E_HsStep.DONE;
        n := 0;
      ELSIF n * GC_CYCLE_MS >= tJob_ms THEN
        xError := TRUE;
        iAlarm := 2;                          (* job time-out *)
      END_IF
    E_HsStep.DONE:
      n := MIN(n + 1, GC_N_MAX);
      IF NOT xDone THEN
        iStep := E_HsStep.IDLE;
        xDoneOut := TRUE;
      ELSIF n * GC_CYCLE_MS >= tHs_ms THEN
        xError := TRUE;
        iAlarm := 3;                          (* done not removed *)
      END_IF
  END_CASE
END_IF
qRequest := (iStep = E_HsStep.REQUEST OR iStep = E_HsStep.BUSY) AND NOT xError;
qEnable := qRequest;
qAck := iStep = E_HsStep.DONE AND NOT xError;
END_FUNCTION_BLOCK

(* ---- FB_Heater.st ---- *)
(*==================================================================================================================
  FB_Heater  -  2-point temperature control with contactor and thermostat monitoring
  ----------------------------------------------------------------------------------------------------------------
  Library   : FMSE device FB library (item 10A)              Version : 1.0.0 (2026-11-15)
  Rule      : tools/fmse/examples/item10a_examples.json  _rules.FB_Heater
  Codegen   : item 8 pattern HEATER -> st_codegen.py calls this FB (x<Signal> / q<Signal>)
  Purpose   : Heater (e.g. washing bath) switched by a contactor: 2-point control with hysteresis below the set
              point, supervision of the contactor feedback (missing / welded), safety thermostat and signal quality.
  Interface :
    dir  name                type          default   meaning
    IN   xOnFb               BOOL          -         contactor auxiliary contact (DI)
    IN   xOverTemp           BOOL          -         safety thermostat tripped (DI)
    IN   rTemp               REAL          20.0      temperature (FB_AnalogIn.rValue)
    IN   xTempGood           BOOL          TRUE      quality GOOD (FB_AnalogIn.xGood)
    IN   xEnable             BOOL          -         heating enabled by the sequence
    IN   rSp                 REAL          60.0      set point
    IN   xReset              BOOL          -         fault reset, rising edge
    CFG  rHyst               REAL          2.0       switch-on hysteresis below rSp
    CFG  tFb_ms              DINT          500       feedback time [ms]
    OUT  qOn                 BOOL          -         heater contactor (DO)
    OUT  xError              BOOL          -         error latched (see alarms)
    OUT  iAlarm              INT           -         local alarm code (0 = none)
  Alarms    : iAlarm = local code a ; Admin.AlarmNo = M*1000 + 10*i + a (decision D2), class per module (D3)
    1  over-temperature (safety thermostat)
    2  no contactor feedback
    3  temperature signal bad
    4  feedback without command (contactor welded?)
  Timing    : Times are counted in calls: n * GC_CYCLE_MS >= t_ms (GC_CYCLE_MS = 100 ms = test bench, TYPES.st).
              In the 10 ms main task set GC_CYCLE_MS := 10 (same behaviour, 10 ms resolution) or replace a counter
              by a TON: ton(IN := <condition>, PT := T#2s); IF ton.Q THEN ... (one call later than the counter).
  Siemens   : SCL (TIA Portal): the same statements; local names are written with '#' (#xRst), the VAR section is
              VAR (STAT) of an FB with an instance DB, R_TRIG / TON are multi-instances, enumerations become INT
              constants (E_DriveState.FAULT -> 9), MIN / LIMIT exist, '16#0080' is written W#16#80 for a WORD.
  NOTICE    : ALL VALUES ARE EXAMPLES. Real PLC code is written, reviewed, tested and signed off by qualified
              people. Safety functions only in the F-program; this FB only reads F-copies and writes no F-signal.
==================================================================================================================*)
FUNCTION_BLOCK FB_Heater
VAR_INPUT  (* signals *)
  xOnFb : BOOL;                             (* contactor auxiliary contact (DI) *)
  xOverTemp : BOOL;                         (* safety thermostat tripped (DI) *)
  rTemp : REAL := 20.0;                     (* temperature (FB_AnalogIn.rValue) *)
  xTempGood : BOOL := TRUE;                 (* quality GOOD (FB_AnalogIn.xGood) *)
  xEnable : BOOL;                           (* heating enabled by the sequence *)
  rSp : REAL := 60.0;                       (* set point *)
  xReset : BOOL;                            (* fault reset, rising edge *)
END_VAR
VAR_INPUT  (* configuration (set once, defaults = example values) *)
  rHyst : REAL := 2.0;                      (* switch-on hysteresis below rSp *)
  tFb_ms : DINT := 500;                     (* feedback time [ms] *)
END_VAR
VAR_OUTPUT  (* outputs *)
  qOn : BOOL;                               (* heater contactor (DO) *)
  xError : BOOL;                            (* error latched (see alarms) *)
  iAlarm : INT;                             (* local alarm code (0 = none) *)
END_VAR
VAR  (* internal *)
  rtReset : R_TRIG;                         (* edge of xReset *)
  xRst : BOOL;                              (* reset pulse *)
  xHeat : BOOL;                             (* 2-point controller state *)
  xQ : BOOL;                                (* contactor command *)
  nFb : DINT;                               (* calls: command without feedback *)
  nWeld : DINT;                             (* calls: feedback without command *)
END_VAR
rtReset(CLK := xReset);
xRst := rtReset.Q;
(* (1) reset only when the cause is gone and the contactor is open *)
IF xError AND xRst AND NOT xOverTemp AND (xTempGood OR NOT xEnable) AND NOT xOnFb THEN
  xError := FALSE;
  iAlarm := 0;
  nFb := 0;
  nWeld := 0;
END_IF
(* (2) thermostat and signal quality *)
IF NOT xError THEN
  IF xOverTemp THEN
    xError := TRUE;
    iAlarm := 1;                              (* over-temperature *)
  ELSIF xEnable AND NOT xTempGood THEN
    xError := TRUE;
    iAlarm := 3;                              (* temperature signal bad *)
  END_IF
END_IF
(* (3) 2-point control: on at rSp - rHyst, off at rSp, unchanged in between *)
IF NOT xEnable OR xError THEN
  xHeat := FALSE;
ELSIF rTemp <= rSp - rHyst THEN
  xHeat := TRUE;
ELSIF rTemp >= rSp THEN
  xHeat := FALSE;
END_IF
xQ := xHeat;
(* (4) contactor feedback supervision *)
IF xQ AND NOT xOnFb THEN
  nFb := MIN(nFb + 1, GC_N_MAX);
ELSE
  nFb := 0;
END_IF
IF NOT xQ AND xOnFb THEN
  nWeld := MIN(nWeld + 1, GC_N_MAX);
ELSE
  nWeld := 0;
END_IF
IF NOT xError AND nFb * GC_CYCLE_MS >= tFb_ms THEN
  xError := TRUE;
  iAlarm := 2;                                (* no contactor feedback *)
END_IF
IF NOT xError AND nWeld * GC_CYCLE_MS >= tFb_ms THEN
  xError := TRUE;
  iAlarm := 4;                                (* feedback without command *)
END_IF
(* (5) an error switches the heater off *)
IF xError THEN
  xHeat := FALSE;
  xQ := FALSE;
END_IF
qOn := xQ;
END_FUNCTION_BLOCK

(* ---- FB_LightCurtain.st ---- *)
(*==================================================================================================================
  FB_LightCurtain  -  light curtain (2 OSSD + warning)
  ----------------------------------------------------------------------------------------------------------------
  Library   : FMSE device FB library (item 10A)              Version : 1.0.0 (2026-11-15)
  Rule      : tools/fmse/examples/item10a_examples.json  _rules.fb_library (= FB_Safe2Ch)
  Codegen   : item 8 pattern LC -> st_codegen.py calls this FB (x<Signal> / q<Signal>)
  Purpose   : Wrapper with the item-8 signal names: xOssd1 / xOssd2 -> FB_Safe2Ch xCh1 / xCh2.
              Diagnosis and HMI only - the safety function is in the F-program.
  Interface :
    dir  name                type          default   meaning
    IN   xOssd1              BOOL          -         OSSD 1 F-copy (TRUE = free)
    IN   xOssd2              BOOL          -         OSSD 2 F-copy (TRUE = free)
    IN   xWarn               BOOL          -         warning / muting signal (DI)
    IN   xReset              BOOL          -         fault reset, rising edge
    CFG  tDisc_ms            DINT          500       discrepancy time [ms]
    OUT  xSafe               BOOL          -         closed / free and reset (FB_Safe2Ch.xOk)
    OUT  xWarnOut            BOOL          -         warning signal passed through
    OUT  xResetReq           BOOL          -         waiting for a reset
    OUT  xDiscErr            BOOL          -         discrepancy latched
    OUT  iAlarm              INT           -         local alarm code (0 = none)
  Alarms    : iAlarm = local code a ; Admin.AlarmNo = M*1000 + 10*i + a (decision D2), class per module (D3)
    1  discrepancy
  Timing    : Times are counted in calls: n * GC_CYCLE_MS >= t_ms (GC_CYCLE_MS = 100 ms = test bench, TYPES.st).
              In the 10 ms main task set GC_CYCLE_MS := 10 (same behaviour, 10 ms resolution) or replace a counter
              by a TON: ton(IN := <condition>, PT := T#2s); IF ton.Q THEN ... (one call later than the counter).
  Siemens   : SCL (TIA Portal): the same statements; local names are written with '#' (#xRst), the VAR section is
              VAR (STAT) of an FB with an instance DB, R_TRIG / TON are multi-instances, enumerations become INT
              constants (E_DriveState.FAULT -> 9), MIN / LIMIT exist, '16#0080' is written W#16#80 for a WORD.
  NOTICE    : ALL VALUES ARE EXAMPLES. Real PLC code is written, reviewed, tested and signed off by qualified
              people. Safety functions only in the F-program; this FB only reads F-copies and writes no F-signal.
==================================================================================================================*)
FUNCTION_BLOCK FB_LightCurtain
VAR_INPUT  (* signals *)
  xOssd1 : BOOL;                            (* OSSD 1 F-copy (TRUE = free) *)
  xOssd2 : BOOL;                            (* OSSD 2 F-copy (TRUE = free) *)
  xWarn : BOOL;                             (* warning / muting signal (DI) *)
  xReset : BOOL;                            (* fault reset, rising edge *)
END_VAR
VAR_INPUT  (* configuration (set once, defaults = example values) *)
  tDisc_ms : DINT := 500;                   (* discrepancy time [ms] *)
END_VAR
VAR_OUTPUT  (* outputs *)
  xSafe : BOOL;                             (* closed / free and reset (FB_Safe2Ch.xOk) *)
  xWarnOut : BOOL;                          (* warning signal passed through *)
  xResetReq : BOOL;                         (* waiting for a reset *)
  xDiscErr : BOOL;                          (* discrepancy latched *)
  iAlarm : INT;                             (* local alarm code (0 = none) *)
END_VAR
VAR  (* internal *)
  fbCh : FB_Safe2Ch;                        (* 2-channel mirror *)
END_VAR
fbCh(xCh1 := xOssd1, xCh2 := xOssd2, xReset := xReset, tDisc_ms := tDisc_ms);
xSafe := fbCh.xOk;
xWarnOut := xWarn;
xResetReq := fbCh.xResetReq;
xDiscErr := fbCh.xDiscErr;
iAlarm := fbCh.iAlarm;
END_FUNCTION_BLOCK

(* ---- FB_LimitAlarm.st ---- *)
(*==================================================================================================================
  FB_LimitAlarm  -  H / L limit alarm with on-delay and hysteresis (item 9)
  ----------------------------------------------------------------------------------------------------------------
  Library   : FMSE device FB library (item 10A)              Version : 1.0.0 (2026-11-15)
  Rule      : tools/fmse/examples/item10a_examples.json  item9_examples.json _rules.limits
  Purpose   : H alarm ON after iDelay consecutive calls with rValue >= rH, OFF at once when rValue < rH - rHyst;
              L alarm ON after iDelay calls with rValue <= rL, OFF when rValue > rL + rHyst.
  Interface :
    dir  name                type          default   meaning
    IN   rValue              REAL          -         process value (FB_AnalogIn.rValue)
    CFG  rH                  REAL          8.0       high limit
    CFG  rL                  REAL          3.0       low limit
    CFG  rHyst               REAL          0.2       hysteresis
    CFG  iDelay              INT           2         on-delay [calls]
    OUT  xH                  BOOL          -         high alarm
    OUT  xL                  BOOL          -         low alarm
  Alarms    : iAlarm = local code a ; Admin.AlarmNo = M*1000 + 10*i + a (decision D2), class per module (D3)
    none
  Timing    : Times are counted in calls: n * GC_CYCLE_MS >= t_ms (GC_CYCLE_MS = 100 ms = test bench, TYPES.st).
              In the 10 ms main task set GC_CYCLE_MS := 10 (same behaviour, 10 ms resolution) or replace a counter
              by a TON: ton(IN := <condition>, PT := T#2s); IF ton.Q THEN ... (one call later than the counter).
  Siemens   : SCL (TIA Portal): the same statements; local names are written with '#' (#xRst), the VAR section is
              VAR (STAT) of an FB with an instance DB, R_TRIG / TON are multi-instances, enumerations become INT
              constants (E_DriveState.FAULT -> 9), MIN / LIMIT exist, '16#0080' is written W#16#80 for a WORD.
  Note      : the counters count CALLS (samples), not milliseconds - one call per sample (item 9: 1 sample/s).
  NOTICE    : ALL VALUES ARE EXAMPLES. Real PLC code is written, reviewed, tested and signed off by qualified
              people. Safety functions only in the F-program; this FB only reads F-copies and writes no F-signal.
==================================================================================================================*)
FUNCTION_BLOCK FB_LimitAlarm
VAR_INPUT  (* signals *)
  rValue : REAL;                            (* process value (FB_AnalogIn.rValue) *)
END_VAR
VAR_INPUT  (* configuration (set once, defaults = example values) *)
  rH : REAL := 8.0;                         (* high limit *)
  rL : REAL := 3.0;                         (* low limit *)
  rHyst : REAL := 0.2;                      (* hysteresis *)
  iDelay : INT := 2;                        (* on-delay [calls] *)
END_VAR
VAR_OUTPUT  (* outputs *)
  xH : BOOL;                                (* high alarm *)
  xL : BOOL;                                (* low alarm *)
END_VAR
VAR  (* internal *)
  nH : DINT;                                (* consecutive calls >= rH *)
  nL : DINT;                                (* consecutive calls <= rL *)
END_VAR
IF rValue >= rH THEN
  nH := MIN(nH + 1, GC_N_MAX);
ELSE
  nH := 0;
END_IF
IF rValue <= rL THEN
  nL := MIN(nL + 1, GC_N_MAX);
ELSE
  nL := 0;
END_IF
IF NOT xH AND nH >= iDelay THEN
  xH := TRUE;
ELSIF xH AND rValue < rH - rHyst THEN
  xH := FALSE;
END_IF
IF NOT xL AND nL >= iDelay THEN
  xL := TRUE;
ELSIF xL AND rValue > rL + rHyst THEN
  xL := FALSE;
END_IF
END_FUNCTION_BLOCK

(* ---- FB_ModeSwitch.st ---- *)
(*==================================================================================================================
  FB_ModeSwitch  -  operating-mode key switch
  ----------------------------------------------------------------------------------------------------------------
  Library   : FMSE device FB library (item 10A)              Version : 1.0.0 (2026-11-15)
  Rule      : tools/fmse/examples/item10a_examples.json  _rules.FB_ModeSwitch
  Codegen   : item 8 pattern MODE_SWITCH -> st_codegen.py calls this FB (x<Signal> / q<Signal>)
  Purpose   : Key switch with two contacts: Auto -> 1 Production, Maint -> 2 Maintenance, none -> 3 Manual;
              both contacts on keeps the last mode and gives an alarm after tDisc_ms.
  Interface :
    dir  name                type          default   meaning
    IN   xAuto               BOOL          -         contact AUTO (DI)
    IN   xMaint              BOOL          -         contact MAINT (DI)
    CFG  tDisc_ms            DINT          500       discrepancy time [ms]
    OUT  iMode               INT           3         1 Production, 2 Maintenance, 3 Manual
    OUT  xError              BOOL          -         error latched (see alarms)
    OUT  iAlarm              INT           -         local alarm code (0 = none)
  Alarms    : iAlarm = local code a ; Admin.AlarmNo = M*1000 + 10*i + a (decision D2), class per module (D3)
    1  both key positions on (discrepancy)
  Timing    : Times are counted in calls: n * GC_CYCLE_MS >= t_ms (GC_CYCLE_MS = 100 ms = test bench, TYPES.st).
              In the 10 ms main task set GC_CYCLE_MS := 10 (same behaviour, 10 ms resolution) or replace a counter
              by a TON: ton(IN := <condition>, PT := T#2s); IF ton.Q THEN ... (one call later than the counter).
  Siemens   : SCL (TIA Portal): the same statements; local names are written with '#' (#xRst), the VAR section is
              VAR (STAT) of an FB with an instance DB, R_TRIG / TON are multi-instances, enumerations become INT
              constants (E_DriveState.FAULT -> 9), MIN / LIMIT exist, '16#0080' is written W#16#80 for a WORD.
  NOTICE    : ALL VALUES ARE EXAMPLES. Real PLC code is written, reviewed, tested and signed off by qualified
              people. Safety functions only in the F-program; this FB only reads F-copies and writes no F-signal.
==================================================================================================================*)
FUNCTION_BLOCK FB_ModeSwitch
VAR_INPUT  (* signals *)
  xAuto : BOOL;                             (* contact AUTO (DI) *)
  xMaint : BOOL;                            (* contact MAINT (DI) *)
END_VAR
VAR_INPUT  (* configuration (set once, defaults = example values) *)
  tDisc_ms : DINT := 500;                   (* discrepancy time [ms] *)
END_VAR
VAR_OUTPUT  (* outputs *)
  iMode : INT := 3;                         (* 1 Production, 2 Maintenance, 3 Manual *)
  xError : BOOL;                            (* error latched (see alarms) *)
  iAlarm : INT;                             (* local alarm code (0 = none) *)
END_VAR
VAR  (* internal *)
  n : DINT;                                 (* calls with both contacts on *)
END_VAR
IF xAuto AND xMaint THEN
  n := MIN(n + 1, GC_N_MAX);
ELSE
  n := 0;
END_IF
IF xAuto AND NOT xMaint THEN
  iMode := E_Mode.PRODUCTION;
ELSIF xMaint AND NOT xAuto THEN
  iMode := E_Mode.MAINTENANCE;
ELSIF NOT xAuto AND NOT xMaint THEN
  iMode := E_Mode.MANUAL;
END_IF                                        (* both on: mode unchanged *)
xError := n * GC_CYCLE_MS >= tDisc_ms;
IF xError THEN
  iAlarm := 1;
ELSE
  iAlarm := 0;
END_IF
END_FUNCTION_BLOCK

(* ---- FB_MotorDol.st ---- *)
(*==================================================================================================================
  FB_MotorDol  -  direct-on-line motor with run-feedback supervision (item 9)
  ----------------------------------------------------------------------------------------------------------------
  Library   : FMSE device FB library (item 10A)              Version : 1.0.0 (2026-11-15)
  Rule      : tools/fmse/examples/item10a_examples.json  item9_examples.json _rules.motor
  Codegen   : item 8 pattern DOL -> st_codegen.py calls this FB (x<Signal> / q<Signal>)
  Purpose   : Contactor motor: start on a rising edge of xCmd (no automatic restart), run feedback after start,
              feedback lost while running, motor protection, feedback without command (welded contactor).
              Reset on a rising edge of xReset only when the cause is gone.
  Interface :
    dir  name                type          default   meaning
    IN   xRunFb              BOOL          -         contactor auxiliary contact (DI)
    IN   xTripped            BOOL          -         motor protection tripped (DI)
    IN   xCmd                BOOL          -         run command from the sequence
    IN   xReset              BOOL          -         fault reset, rising edge
    CFG  tFb_ms              DINT          500       feedback time [ms]
    OUT  qRun                BOOL          -         contactor (DO)
    OUT  iState              INT           -         0 stopped, 1 starting, 2 running, 3 stopping, 9 fault
    OUT  xError              BOOL          -         error latched (see alarms)
    OUT  iAlarm              INT           -         local alarm code (0 = none)
  Alarms    : iAlarm = local code a ; Admin.AlarmNo = M*1000 + 10*i + a (decision D2), class per module (D3)
    1  no run feedback after start
    2  run feedback lost while running
    3  motor protection tripped
    4  run feedback without command (contactor welded?)
  Timing    : Times are counted in calls: n * GC_CYCLE_MS >= t_ms (GC_CYCLE_MS = 100 ms = test bench, TYPES.st).
              In the 10 ms main task set GC_CYCLE_MS := 10 (same behaviour, 10 ms resolution) or replace a counter
              by a TON: ton(IN := <condition>, PT := T#2s); IF ton.Q THEN ... (one call later than the counter).
  Siemens   : SCL (TIA Portal): the same statements; local names are written with '#' (#xRst), the VAR section is
              VAR (STAT) of an FB with an instance DB, R_TRIG / TON are multi-instances, enumerations become INT
              constants (E_DriveState.FAULT -> 9), MIN / LIMIT exist, '16#0080' is written W#16#80 for a WORD.
  NOTICE    : ALL VALUES ARE EXAMPLES. Real PLC code is written, reviewed, tested and signed off by qualified
              people. Safety functions only in the F-program; this FB only reads F-copies and writes no F-signal.
==================================================================================================================*)
FUNCTION_BLOCK FB_MotorDol
VAR_INPUT  (* signals *)
  xRunFb : BOOL;                            (* contactor auxiliary contact (DI) *)
  xTripped : BOOL;                          (* motor protection tripped (DI) *)
  xCmd : BOOL;                              (* run command from the sequence *)
  xReset : BOOL;                            (* fault reset, rising edge *)
END_VAR
VAR_INPUT  (* configuration (set once, defaults = example values) *)
  tFb_ms : DINT := 500;                     (* feedback time [ms] *)
END_VAR
VAR_OUTPUT  (* outputs *)
  qRun : BOOL;                              (* contactor (DO) *)
  iState : INT;                             (* 0 stopped, 1 starting, 2 running, 3 stopping, 9 fault *)
  xError : BOOL;                            (* error latched (see alarms) *)
  iAlarm : INT;                             (* local alarm code (0 = none) *)
END_VAR
VAR  (* internal *)
  rtCmd : R_TRIG;                           (* edge of xCmd *)
  rtReset : R_TRIG;                         (* edge of xReset *)
  n : DINT;                                 (* calls in STARTING / STOPPING *)
  nFb : DINT;                               (* calls with feedback while stopped *)
  xEntered : BOOL;                          (* FAULT entered by the trip in this call *)
END_VAR
rtCmd(CLK := xCmd);
rtReset(CLK := xReset);
xEntered := FALSE;
IF xTripped AND iState <> E_MotorState.FAULT THEN
  iState := E_MotorState.FAULT;
  iAlarm := 3;                                (* motor protection tripped *)
  xEntered := TRUE;
END_IF
IF NOT xEntered THEN
  CASE iState OF
    E_MotorState.STOPPED:
      IF xRunFb THEN
        nFb := MIN(nFb + 1, GC_N_MAX);
      ELSE
        nFb := 0;
      END_IF
      IF nFb * GC_CYCLE_MS >= tFb_ms THEN
        iState := E_MotorState.FAULT;
        iAlarm := 4;                          (* feedback without command *)
      ELSIF rtCmd.Q THEN
        iState := E_MotorState.STARTING;
        n := 0;
      END_IF
    E_MotorState.STARTING:
      n := MIN(n + 1, GC_N_MAX);
      IF xRunFb THEN
        iState := E_MotorState.RUNNING;
      ELSIF n * GC_CYCLE_MS >= tFb_ms THEN
        iState := E_MotorState.FAULT;
        iAlarm := 1;                          (* no run feedback after start *)
      END_IF
    E_MotorState.RUNNING:
      IF NOT xCmd THEN
        iState := E_MotorState.STOPPING;
        n := 0;
      ELSIF NOT xRunFb THEN
        iState := E_MotorState.FAULT;
        iAlarm := 2;                          (* run feedback lost while running *)
      END_IF
    E_MotorState.STOPPING:
      n := MIN(n + 1, GC_N_MAX);
      IF NOT xRunFb THEN
        iState := E_MotorState.STOPPED;
        nFb := 0;
      ELSIF n * GC_CYCLE_MS >= tFb_ms THEN
        iState := E_MotorState.FAULT;
        iAlarm := 4;                          (* feedback without command *)
      END_IF
    E_MotorState.FAULT:
      IF rtReset.Q AND NOT xTripped AND NOT (iAlarm = 4 AND xRunFb) THEN
        iState := E_MotorState.STOPPED;
        iAlarm := 0;
        nFb := 0;
      END_IF
  END_CASE
END_IF
qRun := iState = E_MotorState.STARTING OR iState = E_MotorState.RUNNING;
xError := iState = E_MotorState.FAULT;
END_FUNCTION_BLOCK

(* ---- FB_PushButton.st ---- *)
(*==================================================================================================================
  FB_PushButton  -  illuminated push-button
  ----------------------------------------------------------------------------------------------------------------
  Library   : FMSE device FB library (item 10A)              Version : 1.0.0 (2026-11-15)
  Rule      : tools/fmse/examples/item10a_examples.json  _rules.FB_PushButton
  Codegen   : item 8 pattern PUSHBUTTON -> st_codegen.py calls this FB (x<Signal> / q<Signal>)
  Purpose   : Push-button with lamp: lamp off / on / flashing 1 Hz, pressed level and one-call click pulse.
  Interface :
    dir  name                type          default   meaning
    IN   xPb                 BOOL          -         push-button contact (DI)
    IN   iLampMode           INT           -         0 off, 1 on, 2 flashing
    OUT  qLamp               BOOL          -         lamp (DO)
    OUT  xPressed            BOOL          -         button pressed
    OUT  xClick              BOOL          -         rising edge, one call
  Alarms    : iAlarm = local code a ; Admin.AlarmNo = M*1000 + 10*i + a (decision D2), class per module (D3)
    none
  Timing    : Times are counted in calls: n * GC_CYCLE_MS >= t_ms (GC_CYCLE_MS = 100 ms = test bench, TYPES.st).
              In the 10 ms main task set GC_CYCLE_MS := 10 (same behaviour, 10 ms resolution) or replace a counter
              by a TON: ton(IN := <condition>, PT := T#2s); IF ton.Q THEN ... (one call later than the counter).
  Siemens   : SCL (TIA Portal): the same statements; local names are written with '#' (#xRst), the VAR section is
              VAR (STAT) of an FB with an instance DB, R_TRIG / TON are multi-instances, enumerations become INT
              constants (E_DriveState.FAULT -> 9), MIN / LIMIT exist, '16#0080' is written W#16#80 for a WORD.
  NOTICE    : ALL VALUES ARE EXAMPLES. Real PLC code is written, reviewed, tested and signed off by qualified
              people. Safety functions only in the F-program; this FB only reads F-copies and writes no F-signal.
==================================================================================================================*)
FUNCTION_BLOCK FB_PushButton
VAR_INPUT  (* signals *)
  xPb : BOOL;                               (* push-button contact (DI) *)
  iLampMode : INT;                          (* 0 off, 1 on, 2 flashing *)
END_VAR
VAR_OUTPUT  (* outputs *)
  qLamp : BOOL;                             (* lamp (DO) *)
  xPressed : BOOL;                          (* button pressed *)
  xClick : BOOL;                            (* rising edge, one call *)
END_VAR
VAR  (* internal *)
  nBlink : DINT;                            (* blink counter 0 .. 2*nHalf-1 *)
  nHalf : DINT;                             (* calls per half period *)
  xBlink : BOOL;                            (* 1 Hz blink, TRUE in the first half *)
  rtPb : R_TRIG;                            (* edge of xPb *)
END_VAR
nHalf := GC_BLINK_HALF_MS / GC_CYCLE_MS;     (* 5 calls at 100 ms = 1 Hz *)
xBlink := nBlink < nHalf;
nBlink := (nBlink + 1) MOD (2 * nHalf);
qLamp := (iLampMode = 1) OR ((iLampMode = 2) AND xBlink);
rtPb(CLK := xPb);
xClick := rtPb.Q;
xPressed := xPb;
END_FUNCTION_BLOCK

(* ---- FB_Safe2Ch.st ---- *)
(*==================================================================================================================
  FB_Safe2Ch  -  diagnostic mirror of a 2-channel safety input
  ----------------------------------------------------------------------------------------------------------------
  Library   : FMSE device FB library (item 10A)              Version : 1.0.0 (2026-11-15)
  Rule      : tools/fmse/examples/item10a_examples.json  _rules.FB_Safe2Ch
  Purpose   : Standard-program mirror of a 2-channel safety input (the safety function itself is in the
              F-program): reset needed after power-on and after every opening, discrepancy alarm that can only
              be reset after BOTH channels were open (cross-fault test). Base of FB_Estop, FB_Door2Ch,
              FB_EnableSwitch, FB_LightCurtain and FB_SafetyCoupling.
  Interface :
    dir  name                type          default   meaning
    IN   xCh1                BOOL          -         channel 1, TRUE = safe / closed
    IN   xCh2                BOOL          -         channel 2, TRUE = safe / closed
    IN   xReset              BOOL          -         fault reset, rising edge
    CFG  tDisc_ms            DINT          500       discrepancy time [ms]
    OUT  xOk                 BOOL          -         both channels closed and reset
    OUT  xResetReq           BOOL          -         closed, waiting for a reset (lamp)
    OUT  xDiscErr            BOOL          -         discrepancy latched
    OUT  iAlarm              INT           -         local alarm code (0 = none)
  Alarms    : iAlarm = local code a ; Admin.AlarmNo = M*1000 + 10*i + a (decision D2), class per module (D3)
    1  discrepancy
  Timing    : Times are counted in calls: n * GC_CYCLE_MS >= t_ms (GC_CYCLE_MS = 100 ms = test bench, TYPES.st).
              In the 10 ms main task set GC_CYCLE_MS := 10 (same behaviour, 10 ms resolution) or replace a counter
              by a TON: ton(IN := <condition>, PT := T#2s); IF ton.Q THEN ... (one call later than the counter).
  Siemens   : SCL (TIA Portal): the same statements; local names are written with '#' (#xRst), the VAR section is
              VAR (STAT) of an FB with an instance DB, R_TRIG / TON are multi-instances, enumerations become INT
              constants (E_DriveState.FAULT -> 9), MIN / LIMIT exist, '16#0080' is written W#16#80 for a WORD.
  NOTICE    : ALL VALUES ARE EXAMPLES. Real PLC code is written, reviewed, tested and signed off by qualified
              people. Safety functions only in the F-program; this FB only reads F-copies and writes no F-signal.
==================================================================================================================*)
FUNCTION_BLOCK FB_Safe2Ch
VAR_INPUT  (* signals *)
  xCh1 : BOOL;                              (* channel 1, TRUE = safe / closed *)
  xCh2 : BOOL;                              (* channel 2, TRUE = safe / closed *)
  xReset : BOOL;                            (* fault reset, rising edge *)
END_VAR
VAR_INPUT  (* configuration (set once, defaults = example values) *)
  tDisc_ms : DINT := 500;                   (* discrepancy time [ms] *)
END_VAR
VAR_OUTPUT  (* outputs *)
  xOk : BOOL;                               (* both channels closed and reset *)
  xResetReq : BOOL;                         (* closed, waiting for a reset (lamp) *)
  xDiscErr : BOOL;                          (* discrepancy latched *)
  iAlarm : INT;                             (* local alarm code (0 = none) *)
END_VAR
VAR  (* internal *)
  rtReset : R_TRIG;                         (* edge of xReset *)
  xRst : BOOL;                              (* reset pulse *)
  xLatched : BOOL := TRUE;                  (* reset needed (TRUE after power-on) *)
  nDisc : DINT;                             (* calls with xCh1 <> xCh2 *)
  xBothOpen : BOOL;                         (* both channels were open after the discrepancy *)
END_VAR
rtReset(CLK := xReset);
xRst := rtReset.Q;
IF xCh1 <> xCh2 THEN
  nDisc := MIN(nDisc + 1, GC_N_MAX);
ELSE
  nDisc := 0;
END_IF
IF (nDisc * GC_CYCLE_MS >= tDisc_ms) AND NOT xDiscErr THEN
  xDiscErr := TRUE;
  iAlarm := 1;                                (* discrepancy *)
  xBothOpen := FALSE;
END_IF
IF xDiscErr AND NOT xCh1 AND NOT xCh2 THEN
  xBothOpen := TRUE;
END_IF
IF NOT (xCh1 AND xCh2) THEN
  xLatched := TRUE;
END_IF
IF xRst AND xCh1 AND xCh2 THEN
  IF xDiscErr AND xBothOpen THEN
    xDiscErr := FALSE;
    iAlarm := 0;
  END_IF
  IF NOT xDiscErr THEN
    xLatched := FALSE;
  END_IF
END_IF
xOk := xCh1 AND xCh2 AND NOT xLatched AND NOT xDiscErr;
xResetReq := xLatched AND xCh1 AND xCh2 AND NOT xDiscErr;
END_FUNCTION_BLOCK
